Fanuc KAREL source: kc00015.KL

-- PROVISIONAL review KL for V940-1; original PC SHA256 bef7cca7fd611d85247f53445e4cbee541d75ac21b8b95fc0a8a30e89c9c9fd1
-- Incomplete behavior may be omitted. Consult companion uncertainty JSON. Do not deploy.
PROGRAM KC00015
%NOLOCKGROUP
BEGIN
  -- V9_ZERO_TABLE_METADATA_HINT layout=0002_ascii; no indexed target words; source/name/runtime held
  -- UNRESOLVED_PC offsets 5-12; opcodes 9D,23
  -- UNRESOLVED_PC offsets 17-47; opcodes 27,22,22,27,9D,31,7E,4A
  -- UNRESOLVED_PC offsets 52-56; opcodes 7F
END KC00015
